// TIA Portal V20 export
// export: Created 2026-10-20T12:51:06.4437102Z, ExportSetting WithDefaults, DisplayName Totally Integrated Automation Portal, DisplayVersion V20 Update 6, DisplayName TIA Portal Openness, DisplayVersion V20 Update 6, DisplayName TIA Portal Version Control Interface, DisplayVersion V20 Update 6, DisplayName SINAMICS Startdrive Advanced, DisplayVersion V20 SP1, DisplayName SINAMICS Startdrive G130, G150, S120, S150, SINAMICS MV, G220, S200, S210, DisplayVersion V20 SP1, DisplayName SINAMICS Startdrive G110M, G120, G120C, G120D, G120P, G115D, DisplayVersion V20 SP1, DisplayName STEP 7 Professional, DisplayVersion V20 Update 6, DisplayName STEP 7 Safety, DisplayVersion V20 Update 2, DisplayName WinCC Basic/Comfort/Advanced, DisplayVersion V20 Update 6, DisplayName WinCC Unified, DisplayVersion V20 Update 6
DATA_BLOCK "Main_Panel_DB"   // DB11, F_DB
VERSION : 0.1
// stored: AutoNumber true, DBAccessibleFromOPCUA true, InstanceOfName Main_Panel, InstanceOfType FB
"Main_Panel"
   // VAR_INPUT
   //    Estop_Cabinet_Ch1 : Bool;
   //    Reset_Cabinet : Bool;
   //    Bypass : "F_Bypass_MainPanel";
   // END_VAR
   // VAR_OUTPUT
   //    Safety_OK : Bool;
   //    Main_Panel_OK : Bool;
   //    Bypass_Warning : Bool;
   //    ACK { ExternalAccessible := 'False'; ExternalVisible := 'False'; ExternalWritable := 'False'} : Bool;
   // END_VAR
   // VAR
   //    Estop_Cabinet_DB : ESTOP1;
   // END_VAR
BEGIN
END_DATA_BLOCK
